// Libérer ou remettre à zéro une portée qualité (docs/10 § 10)
{attribute 'pack_mode' := '1'}
TYPE ST_QualityCommand :
STRUCT
    nSeq : UDINT;
    eCmd : E_QualityCmd;
    eScope : E_QualityScope;
    nIndex : USINT;
    nReason : USINT;
    sUser : STRING(24);
END_STRUCT
END_TYPE

(* stored: Version 1.1.0.1, ProductVersion 3.1.4024.12
   DUT ST_QualityCommand: Id {ca4c7be7-77b2-5ca8-aff2-0b8aaeecd119} *)
